// TIA Portal V20 export
// export: Created 2026-10-12T05:14:49.8641043Z, ExportSetting WithDefaults, DisplayName Totally Integrated Automation Portal, DisplayVersion V20, DisplayName TIA Portal Openness, DisplayVersion V20, DisplayName TIA Portal Teamcenter Gateway, DisplayVersion V20, DisplayName TIA Portal Version Control Interface, DisplayVersion V20, DisplayName SINAMICS Startdrive Advanced, DisplayVersion V20 SP1 Update 2, DisplayName SINAMICS Startdrive G110M, G120, G120C, G120D, G120P, G115D, DisplayVersion V20 SP1 Update 2, DisplayName SINAMICS Startdrive G130, G150, S120, S150, SINAMICS MV, G220, S200, S210, DisplayVersion V20 SP1 Update 2, DisplayName STEP 7 Professional, DisplayVersion V20, DisplayName STEP 7 Safety, DisplayVersion V20, DisplayName WinCC Basic/Comfort/Advanced, DisplayVersion V20, DisplayName WinCC Professional, DisplayVersion V20, DisplayName WinCC Unified, DisplayVersion V20
FUNCTION "F_AccessBenchProvision" : Void   // FC168, SCL
{ S7_Optimized_Access := 'TRUE' }
VERSION : 0.1
// stored: AutoNumber true, IsIECCheckEnabled false, SetENOAutomatically false, UDAEnableTagReadback false
BEGIN

   "FRK_LocalUsers".Count := 2;
   "FRK_LocalUsers".Rows[1].User := 'operator';
   "FRK_LocalUsers".Rows[1].Level := 1;
   "FRK_LocalUsers".Rows[1].Salt[0] := BYTE#16#65;
   "FRK_LocalUsers".Rows[1].Salt[1] := BYTE#16#61;
   "FRK_LocalUsers".Rows[1].Salt[2] := BYTE#16#26;
   "FRK_LocalUsers".Rows[1].Salt[3] := BYTE#16#EE;
   "FRK_LocalUsers".Rows[1].Salt[4] := BYTE#16#61;
   "FRK_LocalUsers".Rows[1].Salt[5] := BYTE#16#28;
   "FRK_LocalUsers".Rows[1].Salt[6] := BYTE#16#DF;
   "FRK_LocalUsers".Rows[1].Salt[7] := BYTE#16#A5;
   "FRK_LocalUsers".Rows[1].Salt[8] := BYTE#16#1A;
   "FRK_LocalUsers".Rows[1].Salt[9] := BYTE#16#96;
   "FRK_LocalUsers".Rows[1].Salt[10] := BYTE#16#30;
   "FRK_LocalUsers".Rows[1].Salt[11] := BYTE#16#1C;
   "FRK_LocalUsers".Rows[1].Salt[12] := BYTE#16#C1;
   "FRK_LocalUsers".Rows[1].Salt[13] := BYTE#16#7C;
   "FRK_LocalUsers".Rows[1].Salt[14] := BYTE#16#FF;
   "FRK_LocalUsers".Rows[1].Salt[15] := BYTE#16#32;
   "FRK_LocalUsers".Rows[1].PinHash[0] := BYTE#16#22;
   "FRK_LocalUsers".Rows[1].PinHash[1] := BYTE#16#12;
   "FRK_LocalUsers".Rows[1].PinHash[2] := BYTE#16#AE;
   "FRK_LocalUsers".Rows[1].PinHash[3] := BYTE#16#43;
   "FRK_LocalUsers".Rows[1].PinHash[4] := BYTE#16#35;
   "FRK_LocalUsers".Rows[1].PinHash[5] := BYTE#16#67;
   "FRK_LocalUsers".Rows[1].PinHash[6] := BYTE#16#A3;
   "FRK_LocalUsers".Rows[1].PinHash[7] := BYTE#16#D7;
   "FRK_LocalUsers".Rows[1].PinHash[8] := BYTE#16#C2;
   "FRK_LocalUsers".Rows[1].PinHash[9] := BYTE#16#1C;
   "FRK_LocalUsers".Rows[1].PinHash[10] := BYTE#16#44;
   "FRK_LocalUsers".Rows[1].PinHash[11] := BYTE#16#AE;
   "FRK_LocalUsers".Rows[1].PinHash[12] := BYTE#16#9F;
   "FRK_LocalUsers".Rows[1].PinHash[13] := BYTE#16#22;
   "FRK_LocalUsers".Rows[1].PinHash[14] := BYTE#16#10;
   "FRK_LocalUsers".Rows[1].PinHash[15] := BYTE#16#21;
   "FRK_LocalUsers".Rows[1].PinHash[16] := BYTE#16#59;
   "FRK_LocalUsers".Rows[1].PinHash[17] := BYTE#16#9B;
   "FRK_LocalUsers".Rows[1].PinHash[18] := BYTE#16#24;
   "FRK_LocalUsers".Rows[1].PinHash[19] := BYTE#16#F0;
   "FRK_LocalUsers".Rows[1].PinHash[20] := BYTE#16#A3;
   "FRK_LocalUsers".Rows[1].PinHash[21] := BYTE#16#D2;
   "FRK_LocalUsers".Rows[1].PinHash[22] := BYTE#16#B1;
   "FRK_LocalUsers".Rows[1].PinHash[23] := BYTE#16#DB;
   "FRK_LocalUsers".Rows[1].PinHash[24] := BYTE#16#73;
   "FRK_LocalUsers".Rows[1].PinHash[25] := BYTE#16#59;
   "FRK_LocalUsers".Rows[1].PinHash[26] := BYTE#16#66;
   "FRK_LocalUsers".Rows[1].PinHash[27] := BYTE#16#18;
   "FRK_LocalUsers".Rows[1].PinHash[28] := BYTE#16#FB;
   "FRK_LocalUsers".Rows[1].PinHash[29] := BYTE#16#58;
   "FRK_LocalUsers".Rows[1].PinHash[30] := BYTE#16#9B;
   "FRK_LocalUsers".Rows[1].PinHash[31] := BYTE#16#0C;
   "FRK_LocalUsers".Rows[2].User := 'admin';
   "FRK_LocalUsers".Rows[2].Level := 4;
   "FRK_LocalUsers".Rows[2].Salt[0] := BYTE#16#0E;
   "FRK_LocalUsers".Rows[2].Salt[1] := BYTE#16#A6;
   "FRK_LocalUsers".Rows[2].Salt[2] := BYTE#16#E1;
   "FRK_LocalUsers".Rows[2].Salt[3] := BYTE#16#FF;
   "FRK_LocalUsers".Rows[2].Salt[4] := BYTE#16#A4;
   "FRK_LocalUsers".Rows[2].Salt[5] := BYTE#16#00;
   "FRK_LocalUsers".Rows[2].Salt[6] := BYTE#16#62;
   "FRK_LocalUsers".Rows[2].Salt[7] := BYTE#16#B7;
   "FRK_LocalUsers".Rows[2].Salt[8] := BYTE#16#76;
   "FRK_LocalUsers".Rows[2].Salt[9] := BYTE#16#5F;
   "FRK_LocalUsers".Rows[2].Salt[10] := BYTE#16#8B;
   "FRK_LocalUsers".Rows[2].Salt[11] := BYTE#16#EB;
   "FRK_LocalUsers".Rows[2].Salt[12] := BYTE#16#12;
   "FRK_LocalUsers".Rows[2].Salt[13] := BYTE#16#63;
   "FRK_LocalUsers".Rows[2].Salt[14] := BYTE#16#0A;
   "FRK_LocalUsers".Rows[2].Salt[15] := BYTE#16#F2;
   "FRK_LocalUsers".Rows[2].PinHash[0] := BYTE#16#5D;
   "FRK_LocalUsers".Rows[2].PinHash[1] := BYTE#16#0B;
   "FRK_LocalUsers".Rows[2].PinHash[2] := BYTE#16#5C;
   "FRK_LocalUsers".Rows[2].PinHash[3] := BYTE#16#D5;
   "FRK_LocalUsers".Rows[2].PinHash[4] := BYTE#16#A8;
   "FRK_LocalUsers".Rows[2].PinHash[5] := BYTE#16#43;
   "FRK_LocalUsers".Rows[2].PinHash[6] := BYTE#16#2F;
   "FRK_LocalUsers".Rows[2].PinHash[7] := BYTE#16#86;
   "FRK_LocalUsers".Rows[2].PinHash[8] := BYTE#16#B9;
   "FRK_LocalUsers".Rows[2].PinHash[9] := BYTE#16#89;
   "FRK_LocalUsers".Rows[2].PinHash[10] := BYTE#16#99;
   "FRK_LocalUsers".Rows[2].PinHash[11] := BYTE#16#62;
   "FRK_LocalUsers".Rows[2].PinHash[12] := BYTE#16#95;
   "FRK_LocalUsers".Rows[2].PinHash[13] := BYTE#16#AA;
   "FRK_LocalUsers".Rows[2].PinHash[14] := BYTE#16#01;
   "FRK_LocalUsers".Rows[2].PinHash[15] := BYTE#16#14;
   "FRK_LocalUsers".Rows[2].PinHash[16] := BYTE#16#1E;
   "FRK_LocalUsers".Rows[2].PinHash[17] := BYTE#16#DE;
   "FRK_LocalUsers".Rows[2].PinHash[18] := BYTE#16#6E;
   "FRK_LocalUsers".Rows[2].PinHash[19] := BYTE#16#66;
   "FRK_LocalUsers".Rows[2].PinHash[20] := BYTE#16#3B;
   "FRK_LocalUsers".Rows[2].PinHash[21] := BYTE#16#21;
   "FRK_LocalUsers".Rows[2].PinHash[22] := BYTE#16#3A;
   "FRK_LocalUsers".Rows[2].PinHash[23] := BYTE#16#51;
   "FRK_LocalUsers".Rows[2].PinHash[24] := BYTE#16#A1;
   "FRK_LocalUsers".Rows[2].PinHash[25] := BYTE#16#B8;
   "FRK_LocalUsers".Rows[2].PinHash[26] := BYTE#16#CB;
   "FRK_LocalUsers".Rows[2].PinHash[27] := BYTE#16#5E;
   "FRK_LocalUsers".Rows[2].PinHash[28] := BYTE#16#5D;
   "FRK_LocalUsers".Rows[2].PinHash[29] := BYTE#16#82;
   "FRK_LocalUsers".Rows[2].PinHash[30] := BYTE#16#EA;
   "FRK_LocalUsers".Rows[2].PinHash[31] := BYTE#16#29;

   "GDB_AccessPersistTest".ProvisionCount := "GDB_AccessPersistTest".ProvisionCount + 1;
END_FUNCTION
